# EPICS autosave request: 1.5.0/debian-12/7.0.10/modules/ADCore-ee039d2/db/NDFFT_settings.req
file "NDPluginBase_settings.req", P=$(P), R=$(R)
$(P)$(R)FFTDirection
$(P)$(R)FFTSuppressDC
$(P)$(R)FFTNumAverage
$(P)$(R)Name
